FUNCTION_BLOCK Motor_Inovaisa (* Motor do painel do gradeamento Vibropac (grade ou rosca) - HidrycoLib *)
  (* Standard: 61499-2 *)
  (* Version 1.0, 22/10/2026, Hidryco, Hidryco, 1.0: status de um motor do painel do gradeamento (tabela Modbus Inovaisa PV-35524). IThis com as tags do legado (Grade_Mecanizada_Inovaisa / Motor_Status): STS_FUNCIONAMENTO, STS_SENSOR_SOBRETORQUE, STS_LIGADO, STS_ALARME no evento E_ATUALIZA. Dados pelo processo (sem symlink). *)
  PACKAGE Hidryco.HidrycoLib;
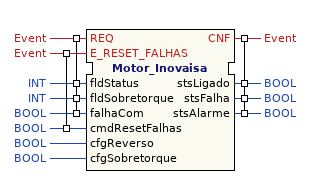
  EVENT_INPUT
    REQ WITH fldStatus, fldSobretorque, falhaCom; (* Leitura do painel (pelo processo) *)
    E_RESET_FALHAS WITH cmdResetFalhas; (* Reconhecimento dos alarmes pelo processo (com cmdResetFalhas = TRUE) *)
  END_EVENT
  EVENT_OUTPUT
    CNF WITH stsLigado, stsFalha, stsAlarme; (* Status (na mudanca) *)
  END_EVENT
  VAR_INPUT
    fldStatus : INT; (* Registro de status do motor (4007/4008/4009) *)
    fldSobretorque : INT; (* Registro do sobretorque (4010/4011) *)
    falhaCom : BOOL; (* Sem comunicacao com o painel *)
    cmdResetFalhas : BOOL; (* TRUE = reconhece (com o evento E_RESET_FALHAS) *)
    cfgReverso : BOOL := FALSE; (* TRUE = grade (avante/reverso); FALSE = rosca *)
    cfgSobretorque : BOOL := FALSE; (* TRUE = tem sensor de sobretorque (grade) *)
  END_VAR
  VAR_OUTPUT
    stsLigado : BOOL; (* Motor funcionando *)
    stsFalha : BOOL; (* Motor em falha *)
    stsAlarme : BOOL; (* Falha ou sobretorque *)
  END_VAR
  FBS
    IThis : Motor_Inovaisa_HMI(QI := TRUE);
    plcStart1 : plcStart(Prio := 10);
    Logica : basicMotorInovaisa;
    AlarmeFalha : ALARM_BIT(TYPE := 1, ACKTYPE_1 := 2, ACTIVE := TRUE); {SET_ATTRIBUTE(HMI.AlarmText, Falha do motor da grade)}
    AlarmeSobretorque : ALARM_BIT(TYPE := 1, ACKTYPE_1 := 2, ACTIVE := TRUE); {SET_ATTRIBUTE(HMI.AlarmText, Sobretorque na grade)}
  END_FBS
  EVENT_CONNECTIONS
    plcStart1.FIRST_INIT TO IThis.ADDA54BBAB97D79C;
    plcStart1.REDO_INIT TO IThis.ADDA54BBAB97D79C;
    IThis.168B52168BE98B03 TO Logica.CC51ED04AC7B8E15;
    REQ TO Logica.1A738D87107B5D6E;
    IThis.2CDECF5265485734 TO Logica.DB88907039BC9764;
    Logica.475E549998D92F9C TO CNF;
    Logica.0DBD7315011AAE6A TO IThis.894CF465CBE5DE99;
    Logica.0DBD7315011AAE6A TO AlarmeFalha.REQ;
    AlarmeFalha.IND_1 TO IThis.894CF465CBE5DE99;
    IThis.2CDECF5265485734 TO AlarmeFalha.ACK_C1;
    E_RESET_FALHAS TO AlarmeFalha.ACK_C1;
    Logica.0DBD7315011AAE6A TO AlarmeSobretorque.REQ;
    AlarmeSobretorque.IND_1 TO IThis.894CF465CBE5DE99;
    IThis.2CDECF5265485734 TO AlarmeSobretorque.ACK_C1;
    E_RESET_FALHAS TO AlarmeSobretorque.ACK_C1;
    Logica.E84D9EC76B90E86C TO AlarmeFalha.INIT;
    AlarmeFalha.INITO TO AlarmeFalha.REQ_INITDATA;
    AlarmeFalha.CNF_INITDATA TO AlarmeFalha.ACTIVATE;
    AlarmeSobretorque.INITO TO AlarmeSobretorque.REQ_INITDATA;
    AlarmeSobretorque.CNF_INITDATA TO AlarmeSobretorque.ACTIVATE;
    AlarmeFalha.INITO TO AlarmeSobretorque.INIT;
    AlarmeSobretorque.INITO TO plcStart1.ACK_FIRST;
  END_CONNECTIONS
  DATA_CONNECTIONS
    cfgReverso TO Logica.2ADC94B6F20E7414;
    cfgSobretorque TO Logica.3FC6EF986F299664;
    fldStatus TO Logica.1CDD71797D6C49E5;
    fldSobretorque TO Logica.7F6C3C59F50BB037;
    falhaCom TO Logica.019BDF7EDEF8F0BD;
    IThis.E70B674576CB02E5 TO Logica.B98B906E7E2460C2;
    Logica.9546553501CAFBCC TO stsLigado;
    Logica.F4944FF8E76D8509 TO stsFalha;
    Logica.33A942412FF6B3E7 TO stsAlarme;
    Logica.24612FD85F48322F TO IThis.F30BD638AF8C13FF;
    Logica.8D8BB9C442BD70AB TO IThis.132A020204BDDA20;
    Logica.9546553501CAFBCC TO IThis.B5F58A52FFB0C024;
    Logica.33A942412FF6B3E7 TO IThis.448B011AAE0077EF;
    Logica.6156601B3E220AA2 TO IThis.F15F28A051648FE4;
    Logica.F4944FF8E76D8509 TO IThis.357502AC3EA2474E;
    Logica.6F41E89DDA623392 TO IThis.84B01C540721AF7B;
    Logica.3A7206A4772B6FAE TO IThis.B43C4E444017CBEB;
    Logica.FB09236565887E17 TO IThis.4360993572C5722B;
    Logica.4B9EC81286BA0C1D TO IThis.0C124BF0C30CD2E9;
    Logica.F4944FF8E76D8509 TO AlarmeFalha.INP;
    AlarmeFalha.STATE_1 TO IThis.ED55F77B30DFA30E;
    Logica.6F41E89DDA623392 TO AlarmeSobretorque.INP;
    AlarmeSobretorque.STATE_1 TO IThis.FF1BB0A2DD9AE219;
  END_CONNECTIONS
END_FUNCTION_BLOCK
